Fanuc KAREL source: ka00080.KL

PROGRAM KA00080
%STACKSIZE=65535
%PRIORITY=65535
%NOLOCKGROUP
VAR
SRC : XYZWPREXT
DST : JOINTPOS9
BEGIN
SRC.X=1.0
-- UNSAFE_SOURCE_IR line 8: DST = convert_xyzwprext_to_jointpos9(SRC)
END KA00080
